FUNCTION FC 1 : INT
BEGIN
END_FUNCTION
